// LIMITA rInput NELL'INTERVALLO [rMinimumValue, rMaximumValue]
FUNCTION F_Saturation : REAL
VAR_INPUT
	rInput			:	REAL;
	rMinimumValue	:	REAL;
	rMaximumValue	:	REAL;
END_VAR
VAR
END_VAR

// ESEGUO UNA SATURAZIONE DEL VALORE IN INGRESSO
F_Saturation	:=	MAX(rMinimumValue, MIN(rMaximumValue, rInput));

END_FUNCTION

(* stored: Version 1.1.0.1, ProductVersion 3.1.4024.9
   POU F_Saturation: Id {c4a9c70a-393f-4194-8b08-98fce22d6591}, SpecialFunc None *)
